// TIA Portal V21 export
TagTable "T_V3"
  X_V3 :   (PLC tag HMI_IF.SwOn, HMI_Connection_1, 100 ms)
